FUNCTION_BLOCK EstocagemLodo (* Estocagem do lodo (900): tanques TQ-01/02 (LIT), sopradores SO-01/02, valvulas VA-01/02 e VB-03/04 - HidrycoLib *)
  (* Standard: 61499-2 *)
  (* Version 1.2, 04/11/2026, Hidryco, Hidryco, 1.2: CNF_NEREDA com H/HH (com tempo, sem memoria) e disponivel dos LIT-900-01/02 para os SludgeHoldingTank1/2 da Nereda; sai na mudanca e a cada 5 s (TickNereda). 1.1: SO sem supervisao de termica (sem sinal no PCE); STP_VEL_SOPRADORES (Hz) no REQ_PARA -> stpVelocidadeAutomatico dos SO. 1.0: divisao da Fase_Solida 1.5 como no legado (estocagem). Sem simbolos proprios: o resumo e os faceplates ficam na DesidratacaoLodo, que recebe CNF_HMI e devolve REQ_PARA, ACK_ALARMES e REQ_EMERG pela camada. *)
  PACKAGE Hidryco.HidrycoLib;
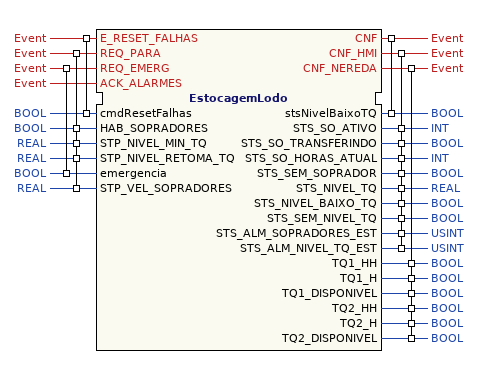
  EVENT_INPUT
    E_RESET_FALHAS WITH cmdResetFalhas; (* Reset pelo processo (estocagem e equipamentos) com cmdResetFalhas = TRUE *)
    REQ_PARA WITH HAB_SOPRADORES, STP_NIVEL_MIN_TQ, STP_NIVEL_RETOMA_TQ, STP_VEL_SOPRADORES; (* DesidratacaoLodo (IHM): ajustes da estocagem *)
    REQ_EMERG WITH emergencia; (* DesidratacaoLodo: emergencia do PCM LODO *)
    ACK_ALARMES; (* DesidratacaoLodo (IHM): reconhecer os alarmes da estocagem *)
  END_EVENT
  EVENT_OUTPUT
    CNF WITH stsNivelBaixoTQ; (* Tanques em nivel baixo (suspende as bombas da DesidratacaoLodo) *)
    CNF_HMI WITH STS_SO_ATIVO, STS_SO_TRANSFERINDO, STS_SO_HORAS_ATUAL, STS_SEM_SOPRADOR, STS_NIVEL_TQ, STS_NIVEL_BAIXO_TQ, STS_SEM_NIVEL_TQ, STS_ALM_SOPRADORES_EST, STS_ALM_NIVEL_TQ_EST; (* Status dos sopradores e tanques para o resumo da DesidratacaoLodo *)
    CNF_NEREDA WITH TQ1_HH, TQ1_H, TQ1_DISPONIVEL, TQ2_HH, TQ2_H, TQ2_DISPONIVEL; (* Nivel dos tanques para a Nereda (SludgeHoldingTank1/2): na mudanca e a cada 5 s *)
  END_EVENT
  VAR_INPUT
    cmdResetFalhas : BOOL; (* TRUE = reset (com o evento E_RESET_FALHAS) *)
    HAB_SOPRADORES : BOOL; (* Da DesidratacaoLodo (IHM): HAB_SOPRADORES *)
    STP_NIVEL_MIN_TQ : REAL; (* Da DesidratacaoLodo (IHM): STP_NIVEL_MIN_TQ *)
    STP_NIVEL_RETOMA_TQ : REAL; (* Da DesidratacaoLodo (IHM): STP_NIVEL_RETOMA_TQ *)
    emergencia : BOOL; (* Emergencia do PCM LODO *)
    STP_VEL_SOPRADORES : REAL := 60.0; (* Da DesidratacaoLodo (IHM): velocidade dos sopradores no automatico (Hz) *)
  END_VAR
  VAR_OUTPUT
    stsNivelBaixoTQ : BOOL; (* Tanques de estocagem em nivel baixo *)
    STS_SO_ATIVO : INT; (* Para a DesidratacaoLodo (IHM): STS_SO_ATIVO *)
    STS_SO_TRANSFERINDO : BOOL; (* Para a DesidratacaoLodo (IHM): STS_SO_TRANSFERINDO *)
    STS_SO_HORAS_ATUAL : INT; (* Para a DesidratacaoLodo (IHM): STS_SO_HORAS_ATUAL *)
    STS_SEM_SOPRADOR : BOOL; (* Para a DesidratacaoLodo (IHM): STS_SEM_SOPRADOR *)
    STS_NIVEL_TQ : REAL; (* Para a DesidratacaoLodo (IHM): STS_NIVEL_TQ *)
    STS_NIVEL_BAIXO_TQ : BOOL; (* Para a DesidratacaoLodo (IHM): STS_NIVEL_BAIXO_TQ *)
    STS_SEM_NIVEL_TQ : BOOL; (* Para a DesidratacaoLodo (IHM): STS_SEM_NIVEL_TQ *)
    STS_ALM_SOPRADORES_EST : USINT; (* Para a DesidratacaoLodo (IHM): STS_ALM_SOPRADORES_EST *)
    STS_ALM_NIVEL_TQ_EST : USINT; (* Para a DesidratacaoLodo (IHM): STS_ALM_NIVEL_TQ_EST *)
    TQ1_HH : BOOL; (* TQ-01 (LIT-900-01): alarme HH com tempo, sem memoria - para o SludgeHoldingTank1 da Nereda *)
    TQ1_H : BOOL; (* TQ-01 (LIT-900-01): alarme H com tempo, sem memoria - para o SludgeHoldingTank1 da Nereda *)
    TQ1_DISPONIVEL : BOOL; (* TQ-01 (LIT-900-01): nivel disponivel (sensor habilitado e sem falha) - para o SludgeHoldingTank1 da Nereda *)
    TQ2_HH : BOOL; (* TQ-02 (LIT-900-02): alarme HH com tempo, sem memoria - para o SludgeHoldingTank2 da Nereda *)
    TQ2_H : BOOL; (* TQ-02 (LIT-900-02): alarme H com tempo, sem memoria - para o SludgeHoldingTank2 da Nereda *)
    TQ2_DISPONIVEL : BOOL; (* TQ-02 (LIT-900-02): nivel disponivel (sensor habilitado e sem falha) - para o SludgeHoldingTank2 da Nereda *)
  END_VAR
  FBS
    IThis : EstocagemLodo_HMI(QI := TRUE);
    plcStart1 : plcStart(Prio := 10);
    Tick : E_CYCLE(DT := T#1s);
    TickNereda : E_CYCLE(DT := T#5s);
    Estocagem : basicEstocagemLodo;
    LIT_900_01 : Sensor_Generico(pin_FC98F78ABCBC0A7E := TRUE, pin_CC8EEC06FF0C4430 := 'm', pin_6D3A2524C5D0F0D1 := 2);
    LIT_900_02 : Sensor_Generico(pin_FC98F78ABCBC0A7E := TRUE, pin_CC8EEC06FF0C4430 := 'm', pin_6D3A2524C5D0F0D1 := 2);
    SO_900_01 : Motor_Generico(pin_D34C88BE7FFF3208 := FALSE, pin_63EFEFB7C85EC93E := TRUE, pin_39489193B7758574 := 600.0);
    SO_900_02 : Motor_Generico(pin_D34C88BE7FFF3208 := FALSE, pin_63EFEFB7C85EC93E := TRUE, pin_39489193B7758574 := 600.0);
    VA_900_01 : Atuador_Coester;
    VA_900_02 : Atuador_Coester;
    VB_900_03 : Atuador_Coester;
    VB_900_04 : Atuador_Coester;
    Revezamento : Controle_Revezamento_2;
    AlarmeSopradores : ALARM_BIT(TYPE := 1, ACKTYPE_1 := 2, ACTIVE := TRUE); {SET_ATTRIBUTE(HMI.AlarmText, Tanques de lodo: nenhum soprador disponível)}
    AlarmeNivelTQ : ALARM_BIT(TYPE := 1, ACKTYPE_1 := 2, ACTIVE := TRUE); {SET_ATTRIBUTE(HMI.AlarmText, Tanques de lodo: nível baixo, bombas suspensas)} {SET_ATTRIBUTE(HMI.AlarmClass, Warning)}
  END_FBS
  EVENT_CONNECTIONS
    AlarmeSopradores.INITO TO AlarmeSopradores.REQ_INITDATA;
    AlarmeSopradores.CNF_INITDATA TO AlarmeSopradores.ACTIVATE;
    AlarmeNivelTQ.INITO TO AlarmeNivelTQ.REQ_INITDATA;
    AlarmeNivelTQ.CNF_INITDATA TO AlarmeNivelTQ.ACTIVATE;
    AlarmeSopradores.INITO TO AlarmeNivelTQ.INIT;
    Tick.EO TO Estocagem.E8C8FA9D941AAB25;
    SO_900_01.9D4F26EE27EDF5B9 TO Estocagem.DFFA20E8FEFD328B;
    Estocagem.A37D04399243417C TO SO_900_01.21070E4B73BFECDC;
    SO_900_02.9D4F26EE27EDF5B9 TO Estocagem.DFFA20E8FEFD328B;
    Estocagem.A37D04399243417C TO SO_900_02.21070E4B73BFECDC;
    LIT_900_01.28A380156DB271B8 TO Estocagem.EA4444D55C79B643;
    LIT_900_02.28A380156DB271B8 TO Estocagem.EA4444D55C79B643;
    REQ_EMERG TO Estocagem.EBAA94C91027AB04;
    Estocagem.820328527C60D44B TO VA_900_01.6AE7937B5439A162;
    Estocagem.820328527C60D44B TO VA_900_02.6AE7937B5439A162;
    Estocagem.820328527C60D44B TO VB_900_03.6AE7937B5439A162;
    Estocagem.820328527C60D44B TO VB_900_04.6AE7937B5439A162;
    REQ_PARA TO Estocagem.C2DAB560DFFB8D5C;
    Estocagem.12E6850BBBD0B68E TO CNF_HMI;
    Estocagem.12E6850BBBD0B68E TO AlarmeSopradores.REQ;
    AlarmeSopradores.IND_1 TO CNF_HMI;
    ACK_ALARMES TO AlarmeSopradores.ACK_C1;
    E_RESET_FALHAS TO AlarmeSopradores.ACK_C1;
    Estocagem.12E6850BBBD0B68E TO AlarmeNivelTQ.REQ;
    AlarmeNivelTQ.IND_1 TO CNF_HMI;
    ACK_ALARMES TO AlarmeNivelTQ.ACK_C1;
    E_RESET_FALHAS TO AlarmeNivelTQ.ACK_C1;
    E_RESET_FALHAS TO LIT_900_01.D21DAA5004F58516;
    E_RESET_FALHAS TO LIT_900_02.D21DAA5004F58516;
    E_RESET_FALHAS TO SO_900_01.BA30A65ADDA4ECC3;
    E_RESET_FALHAS TO SO_900_02.BA30A65ADDA4ECC3;
    E_RESET_FALHAS TO VA_900_01.D903CD18EBE204D1;
    E_RESET_FALHAS TO VA_900_02.D903CD18EBE204D1;
    E_RESET_FALHAS TO VB_900_03.D903CD18EBE204D1;
    E_RESET_FALHAS TO VB_900_04.D903CD18EBE204D1;
    Estocagem.DD4EDADF061294FF TO CNF;
    Revezamento.62818F2F9E2138FC TO Estocagem.C2DAB560DFFB8D5C;
    Estocagem.12E6850BBBD0B68E TO Revezamento.7D54AD64877107DE;
    plcStart1.FIRST_INIT TO IThis.E67C3D572E8F47F1;
    plcStart1.REDO_INIT TO IThis.E67C3D572E8F47F1;
    IThis.F983F3612E0B4890 TO Estocagem.243DC77CA0D0953F;
    Estocagem.5F76B62564497316 TO Tick.START;
    Estocagem.5F76B62564497316 TO Revezamento.1DF068F97CBC55AD;
    Estocagem.5F76B62564497316 TO AlarmeSopradores.INIT;
    AlarmeNivelTQ.INITO TO plcStart1.ACK_FIRST;
    Estocagem.5F76B62564497316 TO TickNereda.START;
    TickNereda.EO TO CNF_NEREDA;
    LIT_900_01.28A380156DB271B8 TO CNF_NEREDA;
    LIT_900_02.28A380156DB271B8 TO CNF_NEREDA;
  END_CONNECTIONS
  DATA_CONNECTIONS
    SO_900_01.EBDC9E59C4286586 TO Estocagem.9D0A018985052F58;
    SO_900_01.40A5976BFB296133 TO Estocagem.C050A723D1972718;
    Estocagem.6EEF3183DA620253 TO SO_900_01.87DAE15414E7C412;
    Estocagem.821D8F0728BFD8D2 TO SO_900_01.85953C7B9294A9BF;
    SO_900_02.EBDC9E59C4286586 TO Estocagem.6442D6171574AD0F;
    SO_900_02.40A5976BFB296133 TO Estocagem.DB889EF87AAB0D82;
    Estocagem.8F8F344FCE172148 TO SO_900_02.87DAE15414E7C412;
    Estocagem.821D8F0728BFD8D2 TO SO_900_02.85953C7B9294A9BF;
    LIT_900_01.E6F78A591442B69F TO Estocagem.76186D6114386881;
    LIT_900_01.726640D1704B3F86 TO Estocagem.DEE813645F20FA9B;
    LIT_900_02.E6F78A591442B69F TO Estocagem.8747D35EC434F184;
    LIT_900_02.726640D1704B3F86 TO Estocagem.284C3EA5513A6D62;
    emergencia TO Estocagem.8603BC9EB66FE144;
    Estocagem.937510DD507F2D1B TO VA_900_01.05903B4B679AA14E;
    Estocagem.937510DD507F2D1B TO VA_900_02.05903B4B679AA14E;
    Estocagem.937510DD507F2D1B TO VB_900_03.05903B4B679AA14E;
    Estocagem.937510DD507F2D1B TO VB_900_04.05903B4B679AA14E;
    HAB_SOPRADORES TO Estocagem.5CF5D34DC0BD4690;
    STP_NIVEL_MIN_TQ TO Estocagem.834BCC8A73E45242;
    STP_NIVEL_RETOMA_TQ TO Estocagem.6A41927EA4F7A44E;
    Estocagem.0C2557554843B422 TO STS_SO_ATIVO;
    Estocagem.0C18C6251210ADD2 TO STS_SO_TRANSFERINDO;
    Estocagem.4235B19D4DDCC680 TO STS_SO_HORAS_ATUAL;
    Estocagem.00131AAE1783E6A4 TO STS_SEM_SOPRADOR;
    Estocagem.27E22A4C9A4D8B67 TO STS_NIVEL_TQ;
    Estocagem.9185345097862782 TO STS_NIVEL_BAIXO_TQ;
    Estocagem.7A648FEA2F2E214A TO STS_SEM_NIVEL_TQ;
    Estocagem.00131AAE1783E6A4 TO AlarmeSopradores.INP;
    AlarmeSopradores.STATE_1 TO STS_ALM_SOPRADORES_EST;
    Estocagem.9185345097862782 TO AlarmeNivelTQ.INP;
    AlarmeNivelTQ.STATE_1 TO STS_ALM_NIVEL_TQ_EST;
    cmdResetFalhas TO LIT_900_01.1908F43CB878F5E7;
    cmdResetFalhas TO LIT_900_02.1908F43CB878F5E7;
    cmdResetFalhas TO SO_900_01.C2F1E9C0FB076F17;
    cmdResetFalhas TO SO_900_02.C2F1E9C0FB076F17;
    cmdResetFalhas TO VA_900_01.C82CBBE25FC56079;
    cmdResetFalhas TO VA_900_02.C82CBBE25FC56079;
    cmdResetFalhas TO VB_900_03.C82CBBE25FC56079;
    cmdResetFalhas TO VB_900_04.C82CBBE25FC56079;
    Estocagem.9185345097862782 TO stsNivelBaixoTQ;
    Revezamento.E20C11B2DD910C9B TO Estocagem.7307922C026394A4;
    Revezamento.8F7C57B973CE6721 TO Estocagem.ABC6D729A9607229;
    Revezamento.B121C963D16B0207 TO Estocagem.F2FB54ACA0B1231D;
    Estocagem.C56DE563E1383C2E TO Revezamento.BCDE1E145B7C7428;
    Estocagem.6097DB009BDB40DE TO Revezamento.B99EA94F80E94BD2;
    Estocagem.53980AC2D919D417 TO Revezamento.30C56EFD8B8A4EB9;
    STP_VEL_SOPRADORES TO Estocagem.AE27A9FC614464FF;
    Estocagem.59B400080C7CCAAB TO SO_900_01.F94ABA993E8E9FF4;
    Estocagem.59B400080C7CCAAB TO SO_900_02.F94ABA993E8E9FF4;
    LIT_900_01.0A7E41873A4DE750 TO TQ1_HH;
    LIT_900_01.41659C068F94B5C6 TO TQ1_H;
    LIT_900_01.B7194E42DC1D5273 TO TQ1_DISPONIVEL;
    LIT_900_02.0A7E41873A4DE750 TO TQ2_HH;
    LIT_900_02.41659C068F94B5C6 TO TQ2_H;
    LIT_900_02.B7194E42DC1D5273 TO TQ2_DISPONIVEL;
  END_CONNECTIONS
END_FUNCTION_BLOCK
